// TIA Portal V20 export
DATA_BLOCK "DataFromSafey_DB"   // DB70
// stored: AssignedProDiagFB ProDiag_Allgemein, InstanceOfName DataFromSafey, InstanceOfType FB
"DataFromSafey"
   // VAR
   //    "Q_NOT-HALT Taster1" : Bool := TRUE;
   //    "Q_NOT-HALT Extern 1" : Bool := TRUE;
   //    "Q_NOT-HALT Extern 2" : Bool := TRUE;
   //    "FDBACK_NOT-HALT Schütz mit DE_NOT-HALT_Schuetz_Rueckf" : Bool := FALSE;
   //    "FDBACK_NOT-HALT Schütz mit IS_Rueck_Entlueftung" : Bool := FALSE;
   //    "FDBACK_NOT-HALT Schütz mit IS_Druckbereich_entlueftet" : Bool := FALSE;
   //    "FDBACK_NOT-HALT Türe 1 RST mit DE_NOT-HALT_Tuere_1_Rueck_RST" : Bool := TRUE;
   //    "FDBACK_NOT-HALT Türe 1 mit DE_NOT-HALT_Tuere_1_Rueckf" : Bool := FALSE;
   //    "FDBACK_NOT-HALT Türe 1 mit DE_Antriebe_Rueckf" : Bool := FALSE;
   //    "FDBACK_NOT-HALT Türe 2 RST mit DE_NOT-HALT_Tuere_2_Rueck_RST" : Bool := TRUE;
   //    "FDBACK_NOT-HALT Türe 2 mit DE_NOT-HALT_Tuere_2_Rueckf" : Bool := TRUE;
   //    "FDBACK_NOT-HALT Schalter OK mit DE_NOT-HALT_Schalter_OK_Rueckf" : Bool;
   // END_VAR
BEGIN
END_DATA_BLOCK
